// TIA Portal V20 export
// export: Created 2026-10-12T16:46:21.5479727Z, ExportSetting WithDefaults, DisplayName Totally Integrated Automation Portal, DisplayVersion V20 Update 6, DisplayName TIA Portal Openness, DisplayVersion V20 Update 6, DisplayName TIA Portal Version Control Interface, DisplayVersion V20 Update 6, DisplayName SINAMICS Startdrive Advanced, DisplayVersion V20 SP1 Update 2, DisplayName SINAMICS Startdrive G110M, G120, G120C, G120D, G120P, G115D, DisplayVersion V20 SP1 Update 2, DisplayName SINAMICS Startdrive G130, G150, S120, S150, SINAMICS MV, G220, S200, S210, DisplayVersion V20 SP1 Update 2, DisplayName STEP 7 Professional, DisplayVersion V20 Update 6, DisplayName STEP 7 Safety, DisplayVersion V20 Update 2, DisplayName WinCC Basic/Comfort/Advanced, DisplayVersion V20 Update 6, DisplayName WinCC Professional, DisplayVersion V20 Update 6, DisplayName WinCC Unified, DisplayVersion V20 Update 6
DATA_BLOCK "DB_Bad_Konfig"   // DB8
{ S7_Optimized_Access := 'TRUE' }
VERSION : 0.5
// stored: AutoNumber true, DBAccessibleFromOPCUA true, DBAccessibleFromWebserver true, IsOnlyStoredInLoadMemory false, IsRetainMemResEnabled false, IsWriteProtectedInAS false, MemoryReserve 100
   VAR
      Bad_Konfig : Array[1.."c_Anzahl_Bad"] of "UDT_Bad_Konfig";
   END_VAR
BEGIN
   Bad_Konfig[7..8].Ausstattung.HatHeizung_1 := TRUE;
   Bad_Konfig[12].Ausstattung.HatHeizung_1 := TRUE;
   Bad_Konfig[25].Ausstattung.HatHeizung_1 := TRUE;
   Bad_Konfig[36].Ausstattung.HatHeizung_1 := TRUE;
   Bad_Konfig[40].Ausstattung.HatHeizung_1 := TRUE;
   Bad_Konfig[46].Ausstattung.HatHeizung_1 := TRUE;
   Bad_Konfig[25].Ausstattung.HatHeizung_2 := TRUE;
   Bad_Konfig[8].Ausstattung.HatPumpe := TRUE;
   Bad_Konfig[12].Ausstattung.HatPumpe := TRUE;
   Bad_Konfig[14].Ausstattung.HatPumpe := TRUE;
   Bad_Konfig[18..19].Ausstattung.HatPumpe := TRUE;
   Bad_Konfig[21].Ausstattung.HatPumpe := TRUE;
   Bad_Konfig[25..26].Ausstattung.HatPumpe := TRUE;
   Bad_Konfig[31].Ausstattung.HatPumpe := TRUE;
   Bad_Konfig[41].Ausstattung.HatPumpe := TRUE;
   Bad_Konfig[45].Ausstattung.HatPumpe := TRUE;
   Bad_Konfig[25].Ausstattung.HatPumpe_FU := TRUE;
   Bad_Konfig[25].Ausstattung.HatWarenbewegung_X := TRUE;
   Bad_Konfig[25].Ausstattung.HatWarenbewegung_Y := TRUE;
   Bad_Konfig[8].Ausstattung.HatUltraschall := TRUE;
   Bad_Konfig[12].Ausstattung.HatUltraschall := TRUE;
   Bad_Konfig[31].Ausstattung.HatGleichrichter := TRUE;
   Bad_Konfig[36].Ausstattung.HatGleichrichter := TRUE;
   Bad_Konfig[40].Ausstattung.HatGleichrichter := TRUE;
   Bad_Konfig[7..8].Ausstattung.HatNiveau := TRUE;
   Bad_Konfig[12].Ausstattung.HatNiveau := TRUE;
   Bad_Konfig[25].Ausstattung.HatNiveau := TRUE;
   Bad_Konfig[36].Ausstattung.HatNiveau := TRUE;
   Bad_Konfig[40].Ausstattung.HatNiveau := TRUE;
   Bad_Konfig[46].Ausstattung.HatNiveau := TRUE;
   Bad_Konfig[1].WT[1..3].Auftragsindex := -1;
   Bad_Konfig[2].WT[1..3].Auftragsindex := -1;
   Bad_Konfig[3].WT[1..3].Auftragsindex := -1;
   Bad_Konfig[4].WT[1..3].Auftragsindex := -1;
   Bad_Konfig[5].WT[1..3].Auftragsindex := -1;
   Bad_Konfig[6].WT[1..3].Auftragsindex := -1;
   Bad_Konfig[7].WT[1..3].Auftragsindex := -1;
   Bad_Konfig[8].WT[1..3].Auftragsindex := -1;
   Bad_Konfig[9].WT[1..3].Auftragsindex := -1;
   Bad_Konfig[10].WT[1..3].Auftragsindex := -1;
   Bad_Konfig[11].WT[1..3].Auftragsindex := -1;
   Bad_Konfig[12].WT[1..3].Auftragsindex := -1;
   Bad_Konfig[13].WT[1..3].Auftragsindex := -1;
   Bad_Konfig[14].WT[1..3].Auftragsindex := -1;
   Bad_Konfig[15].WT[1..3].Auftragsindex := -1;
   Bad_Konfig[16].WT[1..3].Auftragsindex := -1;
   Bad_Konfig[17].WT[1..3].Auftragsindex := -1;
   Bad_Konfig[18].WT[1..3].Auftragsindex := -1;
   Bad_Konfig[19].WT[1..3].Auftragsindex := -1;
   Bad_Konfig[20].WT[1..3].Auftragsindex := -1;
   Bad_Konfig[21].WT[1..3].Auftragsindex := -1;
   Bad_Konfig[22].WT[1..3].Auftragsindex := -1;
   Bad_Konfig[23].WT[1..3].Auftragsindex := -1;
   Bad_Konfig[24].WT[1..3].Auftragsindex := -1;
   Bad_Konfig[25].WT[1..3].Auftragsindex := -1;
   Bad_Konfig[26].WT[1..3].Auftragsindex := -1;
   Bad_Konfig[27].WT[1..3].Auftragsindex := -1;
   Bad_Konfig[28].WT[1..3].Auftragsindex := -1;
   Bad_Konfig[29].WT[1..3].Auftragsindex := -1;
   Bad_Konfig[30].WT[1..3].Auftragsindex := -1;
   Bad_Konfig[31].WT[1..3].Auftragsindex := -1;
   Bad_Konfig[32].WT[1..3].Auftragsindex := -1;
   Bad_Konfig[33].WT[1..3].Auftragsindex := -1;
   Bad_Konfig[34].WT[1..3].Auftragsindex := -1;
   Bad_Konfig[35].WT[1..3].Auftragsindex := -1;
   Bad_Konfig[36].WT[1..3].Auftragsindex := -1;
   Bad_Konfig[37].WT[1..3].Auftragsindex := -1;
   Bad_Konfig[38].WT[1..3].Auftragsindex := -1;
   Bad_Konfig[39].WT[1..3].Auftragsindex := -1;
   Bad_Konfig[40].WT[1..3].Auftragsindex := -1;
   Bad_Konfig[41].WT[1..3].Auftragsindex := -1;
   Bad_Konfig[42].WT[1..3].Auftragsindex := -1;
   Bad_Konfig[43].WT[1..3].Auftragsindex := -1;
   Bad_Konfig[44].WT[1..3].Auftragsindex := -1;
   Bad_Konfig[45].WT[1..3].Auftragsindex := -1;
   Bad_Konfig[46].WT[1..3].Auftragsindex := -1;
   Bad_Konfig[47].WT[1..3].Auftragsindex := -1;
   Bad_Konfig[1].WT[1..3].SchrittIndex := -1;
   Bad_Konfig[2].WT[1..3].SchrittIndex := -1;
   Bad_Konfig[3].WT[1..3].SchrittIndex := -1;
   Bad_Konfig[4].WT[1..3].SchrittIndex := -1;
   Bad_Konfig[5].WT[1..3].SchrittIndex := -1;
   Bad_Konfig[6].WT[1..3].SchrittIndex := -1;
   Bad_Konfig[7].WT[1..3].SchrittIndex := -1;
   Bad_Konfig[8].WT[1..3].SchrittIndex := -1;
   Bad_Konfig[9].WT[1..3].SchrittIndex := -1;
   Bad_Konfig[10].WT[1..3].SchrittIndex := -1;
   Bad_Konfig[11].WT[1..3].SchrittIndex := -1;
   Bad_Konfig[12].WT[1..3].SchrittIndex := -1;
   Bad_Konfig[13].WT[1..3].SchrittIndex := -1;
   Bad_Konfig[14].WT[1..3].SchrittIndex := -1;
   Bad_Konfig[15].WT[1..3].SchrittIndex := -1;
   Bad_Konfig[16].WT[1..3].SchrittIndex := -1;
   Bad_Konfig[17].WT[1..3].SchrittIndex := -1;
   Bad_Konfig[18].WT[1..3].SchrittIndex := -1;
   Bad_Konfig[19].WT[1..3].SchrittIndex := -1;
   Bad_Konfig[20].WT[1..3].SchrittIndex := -1;
   Bad_Konfig[21].WT[1..3].SchrittIndex := -1;
   Bad_Konfig[22].WT[1..3].SchrittIndex := -1;
   Bad_Konfig[23].WT[1..3].SchrittIndex := -1;
   Bad_Konfig[24].WT[1..3].SchrittIndex := -1;
   Bad_Konfig[25].WT[1..3].SchrittIndex := -1;
   Bad_Konfig[26].WT[1..3].SchrittIndex := -1;
   Bad_Konfig[27].WT[1..3].SchrittIndex := -1;
   Bad_Konfig[28].WT[1..3].SchrittIndex := -1;
   Bad_Konfig[29].WT[1..3].SchrittIndex := -1;
   Bad_Konfig[30].WT[1..3].SchrittIndex := -1;
   Bad_Konfig[31].WT[1..3].SchrittIndex := -1;
   Bad_Konfig[32].WT[1..3].SchrittIndex := -1;
   Bad_Konfig[33].WT[1..3].SchrittIndex := -1;
   Bad_Konfig[34].WT[1..3].SchrittIndex := -1;
   Bad_Konfig[35].WT[1..3].SchrittIndex := -1;
   Bad_Konfig[36].WT[1..3].SchrittIndex := -1;
   Bad_Konfig[37].WT[1..3].SchrittIndex := -1;
   Bad_Konfig[38].WT[1..3].SchrittIndex := -1;
   Bad_Konfig[39].WT[1..3].SchrittIndex := -1;
   Bad_Konfig[40].WT[1..3].SchrittIndex := -1;
   Bad_Konfig[41].WT[1..3].SchrittIndex := -1;
   Bad_Konfig[42].WT[1..3].SchrittIndex := -1;
   Bad_Konfig[43].WT[1..3].SchrittIndex := -1;
   Bad_Konfig[44].WT[1..3].SchrittIndex := -1;
   Bad_Konfig[45].WT[1..3].SchrittIndex := -1;
   Bad_Konfig[46].WT[1..3].SchrittIndex := -1;
   Bad_Konfig[47].WT[1..3].SchrittIndex := -1;
END_DATA_BLOCK
